(* IEC 61131-3 sources: kns-port-domestic/tools/port_metrics_tests/fixtures/adapted/src/POUs/F_Scale, 2 files *)

(* ---- F_Scale.decl.st ---- *)
FUNCTION F_Scale : REAL
VAR_INPUT
    rIn : REAL;
    rK : REAL;
END_VAR

(* ---- F_Scale.impl.st ---- *)
F_Scale := rIn * rK;
IF rK = 0.0 THEN
    F_Scale := 0.0;
END_IF
// PORT: [build] ограничение вынесено в вызывающий код (docs/BUILD_ERRORS.md, запись 1)
